ABB RAPID module: SplitP.mod

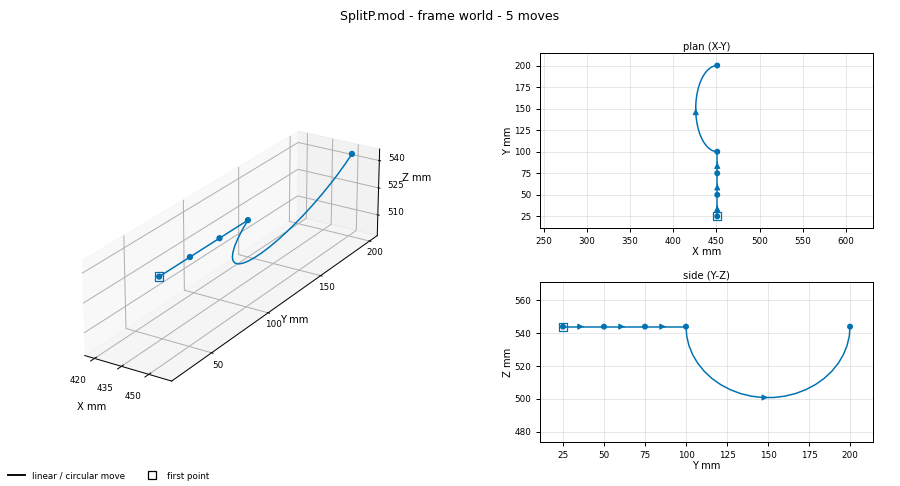
[picture p0: tool path of SplitP.mod in frame world, 5 of 6 moves have a stored position in this frame; points joined in program order, loops and branches not executed]
%%%
  VERSION:1
  LANGUAGE:ENGLISH
%%%
MODULE MOD_SplitP

    ! -------------------------------
    ! Define customized variables here
    ! ...

	! Tool variables:
	PERS tooldata T1 := [TRUE,[[0.000,0.000,100.000],[1.00000000,0.00000000,0.00000000,0.00000000]],[1,[0,0,20],[1,0,0,0],0,0,0.005]];

	! Reference variables:
	PERS wobjdata F1 := [FALSE, TRUE, "", [[0,0,0],[1,0,0,0]],[[0.000,1000.000,0.000],[1.00000000,0.00000000,0.00000000,0.00000000]]];

	PROC Main()
		ConfJ \On;
		ConfL \Off;
		! Program generated by RoboDK v6.0.7 for ABB IRB 120-3/0.6 on XX/XX/XXXX 13:14:16
		! Using nominal kinematics.
		MoveAbsJ [[0.000000,0.000000,0.000000,0.000000,30.000000,-0.000000],[9E+09,9E+09,9E+09,9E+09,9E+09,9E+09]],v500,z1,T1 \WObj:=F1;
		! Splitting Linear movement in 4 (instruction 3: MoveL (S1))
		MoveL [[450.956,-975.000,544.000],[0.50000000,-0.00000001,0.86602540,0.00000000],[0,-1,0,0],[9E+09,9E+09,9E+09,9E+09,9E+09,9E+09]],v500,z1,T1 \WObj:=F1;
		MoveL [[450.956,-950.000,544.000],[0.50000000,-0.00000001,0.86602540,0.00000000],[0,-1,0,0],[9E+09,9E+09,9E+09,9E+09,9E+09,9E+09]],v500,z1,T1 \WObj:=F1;
		MoveL [[450.956,-925.000,544.000],[0.50000000,-0.00000001,0.86602540,-0.00000000],[0,-1,0,0],[9E+09,9E+09,9E+09,9E+09,9E+09,9E+09]],v500,z1,T1 \WObj:=F1;
		MoveL [[450.956,-900.000,544.000],[0.50000000,-0.00000001,0.86602540,-0.00000000],[0,-1,0,0],[9E+09,9E+09,9E+09,9E+09,9E+09,9E+09]],v500,z1,T1 \WObj:=F1;
		MoveC [[425.956,-850.000,500.699],[0.50000000,-0.00000001,0.86602540,-0.00000000],[0,0,-1,0],[9E+09,9E+09,9E+09,9E+09,9E+09,9E+09]],[[450.956,-800.000,544.000],[0.50000000,-0.00000001,0.86602540,-0.00000000],[0,0,-1,0],[9E+09,9E+09,9E+09,9E+09,9E+09,9E+09]],v500,z1,T1 \WObj:=F1;
	ENDPROC

ENDMODULE
